FUNCTION_BLOCK FB_BOSCHINDRADRIVECIA402_REF
VAR_INPUT
	lrScalingFactor 		:LREAL;						(* Position scaling factor *)	
	
	bDriverZKL3				:BOOL;						(* Drive change bit class 3 diagnostics *)
	bDriverZKL2				:BOOL;						(* Drive change bit class 2 diagnostics *)
	bDriverZKL1				:BOOL;						(* Drive error, error in class 1 diagnostics *)
	
	bDriveBB				:BOOL;						(* Drive ready for power on *)
	bDriveAB				:BOOL;						(* Drive control section and power section ready for operation, torque-free*)
	bDriveAF				:BOOL;						(* Drive in operation, with torque *)	
	
	stTerminalState			AT %I*:ST_TerminalState;
	stBoschToPlc			AT %I*:ST_BOSCHINDRADRIVECIA402TOPLC;
	stPlcToBosch			AT %Q*:ST_PLCTOBOSCHINDRADRIVECIA402;
END_VAR
VAR_OUTPUT
	
END_VAR
VAR
	
END_VAR


;

END_FUNCTION_BLOCK

(* stored: Version 1.1.0.1, ProductVersion 3.1.4024.15
   POU FB_BOSCHINDRADRIVECIA402_REF: Id {173232fa-9edf-4c12-82f4-c84611207772}, SpecialFunc None *)
